(* PLC project case, CODESYS CODESYS V3.5 SP17 Patch 3 *)
(* stored: creationDateTime 2026-10-20T00:00:00 *)

CONFIGURATION Device
  RESOURCE Application ON PLC
  END_RESOURCE
END_CONFIGURATION

CONFIGURATION Watchdog
END_CONFIGURATION
